(* IEC 61131-3 sources: KinematicsSimulation/crates/sim-opcua/examples/plc/codesys, 3 files *)

(* ---- sim_cycle.st ---- *)
(*
    A PLC cycle against the KinematicsSimulation link (sim-opcua), for CODESYS V3.5 with the CODESYS OPC UA Client
    SL (PLCopen "OPC UA Client for IEC 61131-3" blocks). Uses SIM_Access, SIM_MC_Power and SIM_MC_MoveAbsolute from
    sim_plcopen.st in this folder.

    NOT COMPILED: CODESYS needs a CODESYS Store account to download, so it was not built. The names follow the
    PLCopen specification OPC 30001 (PLCopen-CFB) v1.02, checked 14 November 2026 at reference.opcfoundation.org.
    CHECK: CODESYS's public help shows only its object-oriented "OPC UA Client" library (Client, Read, Write, ...),
    not these PLCopen blocks; a library that offers them may need its namespace prefix. Spec v1.02 also lists
    UA_NamespaceGetIndex, UA_NodeGetHandle, UA_Read and UA_Write as phased out in favour of their *List variants.

    PRG_SimCycle does what ../twincat/sim_cycle.st does: connect with Basic256Sha256 SignAndEncrypt (or None) and
    optionally user name and password, find the namespace index, power the axis, MC_MoveAbsolute, write a path and
    run it, wait until status.busy falls, switch off and disconnect; meanwhile it reads the axis position and
    following error every cycle through node handles got once. Run it in a task of 10 ms.

    Data types (docs/plc.md, "Node ids and data types"): Double -> LREAL, Boolean -> BOOL, UInt16 -> UINT,
    Int32 -> DINT, UInt64 -> ULINT, String -> STRING. The value of UA_Read/UA_Write is an IN_OUT of type ANY: its
    IEC type is what goes on the wire, so it has to be the one in the table.
*)

FUNCTION_BLOCK SIM_CyclicRead
(* Reads one LREAL variable over and over through a node handle that is got once. *)
VAR_INPUT
    xEnable     : BOOL;
    hConnection : DWORD;
    uiNamespace : UINT;
    sNode       : STRING(255);
END_VAR
VAR_OUTPUT
    lrValue   : LREAL;
    udiReads  : UDINT;
    xError    : BOOL;
    dwErrorID : DWORD;
END_VAR
VAR
    fbGetHandle : UA_NodeGetHandle;
    fbRead      : UA_Read;
    fbRelease   : UA_NodeReleaseHandle;
    stNodeID    : UANodeID;
    stInfo      : UANodeAdditionalInfo;
    hNode       : DWORD;
    iStep       : INT;
END_VAR

CASE iStep OF
0:  IF xEnable THEN
        stNodeID.NamespaceIndex := uiNamespace;
        stNodeID.Identifier := sNode;
        stNodeID.IdentifierType := UAIdentifierType.UAIT_String;
        stInfo.AttributeID := 13;   (* the Value attribute *)
        xError := FALSE; dwErrorID := 0;
        iStep := 1;
    END_IF
1:  fbGetHandle(Execute := TRUE, ConnectionHdl := hConnection, NodeID := stNodeID, Timeout := T#5S);
    IF fbGetHandle.Done THEN
        hNode := fbGetHandle.NodeHdl; fbGetHandle(Execute := FALSE, ConnectionHdl := hConnection, NodeID := stNodeID);
        iStep := 2;
    ELSIF fbGetHandle.Error THEN
        dwErrorID := fbGetHandle.ErrorID; fbGetHandle(Execute := FALSE, ConnectionHdl := hConnection, NodeID := stNodeID);
        xError := TRUE; iStep := 9;
    END_IF
2:  (* once a read is done the next starts in the same cycle *)
    fbRead(Execute := TRUE, ConnectionHdl := hConnection, NodeHdl := hNode, NodeAddInfo := stInfo, Timeout := T#5S,
           Variable := lrValue);
    IF fbRead.Done OR fbRead.Error THEN
        IF fbRead.Error THEN xError := TRUE; dwErrorID := fbRead.ErrorID; ELSE udiReads := udiReads + 1; END_IF
        fbRead(Execute := FALSE, Variable := lrValue);
        IF xEnable THEN
            fbRead(Execute := TRUE, ConnectionHdl := hConnection, NodeHdl := hNode, NodeAddInfo := stInfo,
                   Timeout := T#5S, Variable := lrValue);
        ELSE
            iStep := 3;
        END_IF
    END_IF
3:  fbRelease(Execute := TRUE, ConnectionHdl := hConnection, NodeHdl := hNode, Timeout := T#5S);
    IF fbRelease.Done OR fbRelease.Error THEN
        fbRelease(Execute := FALSE, ConnectionHdl := hConnection, NodeHdl := hNode); iStep := 0;
    END_IF
9:  IF NOT xEnable THEN iStep := 0; END_IF
END_CASE
END_FUNCTION_BLOCK

FUNCTION_BLOCK SIM_WriteString
(* One write of a STRING variable: get the handle, write, release. *)
VAR_INPUT
    xExecute    : BOOL;
    hConnection : DWORD;
    uiNamespace : UINT;
    sNode       : STRING(255);
END_VAR
VAR_IN_OUT
    sValue : STRING(255);
END_VAR
VAR_OUTPUT
    xDone : BOOL; xError : BOOL; dwErrorID : DWORD;
END_VAR
VAR
    fbGetHandle : UA_NodeGetHandle;
    fbWrite     : UA_Write;
    fbRelease   : UA_NodeReleaseHandle;
    stNodeID    : UANodeID;
    stInfo      : UANodeAdditionalInfo;
    hNode       : DWORD;
    iStep       : INT;
    xLast       : BOOL;
END_VAR

IF xExecute AND NOT xLast THEN
    xDone := FALSE; xError := FALSE; dwErrorID := 0;
    stNodeID.NamespaceIndex := uiNamespace;
    stNodeID.Identifier := sNode;
    stNodeID.IdentifierType := UAIdentifierType.UAIT_String;
    stInfo.AttributeID := 13;
    iStep := 1;
END_IF
xLast := xExecute;

CASE iStep OF
1:  fbGetHandle(Execute := TRUE, ConnectionHdl := hConnection, NodeID := stNodeID, Timeout := T#5S);
    IF fbGetHandle.Done THEN
        hNode := fbGetHandle.NodeHdl; fbGetHandle(Execute := FALSE, ConnectionHdl := hConnection, NodeID := stNodeID);
        iStep := 2;
    ELSIF fbGetHandle.Error THEN
        dwErrorID := fbGetHandle.ErrorID; fbGetHandle(Execute := FALSE, ConnectionHdl := hConnection, NodeID := stNodeID);
        xError := TRUE; iStep := 0;
    END_IF
2:  fbWrite(Execute := TRUE, ConnectionHdl := hConnection, NodeHdl := hNode, NodeAddInfo := stInfo, Timeout := T#5S,
            Variable := sValue);
    IF fbWrite.Done OR fbWrite.Error THEN
        xError := fbWrite.Error; dwErrorID := fbWrite.ErrorID;
        fbWrite(Execute := FALSE, Variable := sValue);
        iStep := 3;
    END_IF
3:  fbRelease(Execute := TRUE, ConnectionHdl := hConnection, NodeHdl := hNode, Timeout := T#5S);
    IF fbRelease.Done OR fbRelease.Error THEN
        fbRelease(Execute := FALSE, ConnectionHdl := hConnection, NodeHdl := hNode);
        xDone := NOT xError; iStep := 0;
    END_IF
END_CASE
END_FUNCTION_BLOCK

PROGRAM PRG_SimCycle
VAR
    sServerUrl   : STRING(255) := 'opc.tcp://127.0.0.1:4840';   (* sim-opcua on the same PC *)
    xSecure      : BOOL := TRUE;                                 (* FALSE: SecurityPolicy None *)
    sUser        : STRING(63) := '';                             (* empty: anonymous; else as sim-opcua --user *)
    sPassword    : STRING(63) := '';
    sAxis        : STRING(31) := 'x';
    lrTarget     : LREAL := 0.4;
    sPath        : STRING(255) := 'line,0.4,0.25$Nline,0.1,0.25$Nline,0.1,0.35';
    (* FALSE: the position alone, one Read request a cycle, so that status.client_read_* show the task's cycle *)
    xReadFollowingError : BOOL := TRUE;

    fbConnect    : UA_Connect;
    fbNamespace  : UA_NamespaceGetIndex;
    fbDisconnect : UA_Disconnect;
    stSession    : UASessionConnectInfo;
    hConnection  : DWORD;
    uiNamespace  : UINT;
    fbPower      : SIM_MC_Power;
    fbMove       : SIM_MC_MoveAbsolute;
    fbPath       : SIM_WriteString;
    fbAccess     : SIM_Access;
    fbPosition   : SIM_CyclicRead;
    fbError      : SIM_CyclicRead;
    xFlag        : BOOL;
    lrUnused     : LREAL;
    uiUnused     : UINT;
    xBusySeen    : BOOL;
    lrLargestError : LREAL;
    iStep        : INT;
END_VAR

CASE iStep OF
0:  stSession.ApplicationName := 'CODESYS sim client';
    IF xSecure THEN
        (* The client certificate: create it in View > Security Screen, Devices tab, for the device. sim-opcua
           refuses it once and stores it in pki/rejected; move it to pki/trusted, or run sim-opcua with --trust-all
           while commissioning. The server's certificate (pki/own/cert.der) lands in the device's "Certificates in
           Quarantine" on the first attempt: drag it to "Trusted Certificates" in the same tab. *)
        stSession.SecurityMsgMode := UASecurityMsgMode.UASMM_SignEncrypt;
        stSession.SecurityPolicy := UASecurityPolicy.UASP_Basic256Sha256;
    ELSE
        stSession.SecurityMsgMode := UASecurityMsgMode.UASMM_None;
        stSession.SecurityPolicy := UASecurityPolicy.UASP_None;
    END_IF
    IF LEN(sUser) > 0 THEN
        stSession.UserIdentityToken.UserIdentityTokenType := UAUserIdentityTokenType.UAUITT_Username;
        stSession.UserIdentityToken.TokenParam1 := sUser;
        stSession.UserIdentityToken.TokenParam2 := sPassword;
    END_IF
    fbConnect(Execute := TRUE, ServerEndpointUrl := sServerUrl, SessionConnectInfo := stSession, Timeout := T#5S);
    IF fbConnect.Done THEN hConnection := fbConnect.ConnectionHdl; fbConnect(Execute := FALSE); iStep := 10;
    ELSIF fbConnect.Error THEN fbConnect(Execute := FALSE); iStep := 900; END_IF
10: fbNamespace(Execute := TRUE, ConnectionHdl := hConnection, NamespaceUri := 'urn:kinematics-simulation', Timeout := T#5S);
    IF fbNamespace.Done THEN uiNamespace := fbNamespace.NamespaceIndex; fbNamespace(Execute := FALSE); iStep := 20;
    ELSIF fbNamespace.Error THEN fbNamespace(Execute := FALSE); iStep := 900; END_IF
20: fbPower.Enable := TRUE;
    IF fbPower.Status THEN iStep := 30; END_IF
30: fbMove.Position := lrTarget; fbMove.Velocity := 0.5; fbMove.Acceleration := 5.0; fbMove.Deceleration := 5.0;
    fbMove.Jerk := 100.0;
    fbMove.Execute := TRUE;
    IF fbMove.Done THEN fbMove.Execute := FALSE; iStep := 40;
    ELSIF fbMove.Error OR fbMove.CommandAborted THEN iStep := 900; END_IF
40: fbPath(xExecute := FALSE, sValue := sPath);
    fbPath(xExecute := TRUE, hConnection := hConnection, uiNamespace := uiNamespace, sNode := 'command.path', sValue := sPath);
    IF fbPath.xDone THEN iStep := 42; ELSIF fbPath.xError THEN iStep := 900; ELSE iStep := 41; END_IF
41: fbPath(xExecute := TRUE, sValue := sPath);
    IF fbPath.xDone THEN iStep := 42; ELSIF fbPath.xError THEN iStep := 900; END_IF
42: xFlag := TRUE;
    fbAccess(xExecute := FALSE, xValue := xFlag, lrValue := lrUnused, uiValue := uiUnused);
    fbAccess(xExecute := TRUE, hConnection := hConnection, uiNamespace := uiNamespace, sNode := 'command.run_path',
             eKind := SIM_BOOL, xWrite := TRUE, xValue := xFlag, lrValue := lrUnused, uiValue := uiUnused);
    iStep := 43;
43: fbAccess(xExecute := TRUE, xValue := xFlag, lrValue := lrUnused, uiValue := uiUnused);
    IF fbAccess.xDone THEN xBusySeen := FALSE; iStep := 50; ELSIF fbAccess.xError THEN iStep := 900; END_IF
50: (* poll status.busy until the path is over *)
    fbAccess(xExecute := FALSE, xValue := xFlag, lrValue := lrUnused, uiValue := uiUnused);
    fbAccess(xExecute := TRUE, hConnection := hConnection, uiNamespace := uiNamespace, sNode := 'status.busy',
             eKind := SIM_BOOL, xWrite := FALSE, xValue := xFlag, lrValue := lrUnused, uiValue := uiUnused);
    iStep := 51;
51: fbAccess(xExecute := TRUE, xValue := xFlag, lrValue := lrUnused, uiValue := uiUnused);
    IF fbAccess.xDone THEN
        IF xFlag THEN xBusySeen := TRUE; iStep := 50;
        ELSIF xBusySeen THEN iStep := 60;
        ELSE iStep := 50; END_IF
    ELSIF fbAccess.xError THEN iStep := 900; END_IF
60: fbPower.Enable := FALSE;
    IF NOT fbPower.Status THEN iStep := 70; END_IF
70: fbDisconnect(Execute := TRUE, ConnectionHdl := hConnection, Timeout := T#5S);
    IF fbDisconnect.Done OR fbDisconnect.Error THEN fbDisconnect(Execute := FALSE); iStep := 100; END_IF
100: ; (* finished: lrLargestError holds the largest following error *)
900: ; (* error: look at the blocks' ErrorID and at status.refused on the server *)
END_CASE

fbPosition(xEnable := iStep >= 20 AND iStep < 70, hConnection := hConnection, uiNamespace := uiNamespace,
           sNode := CONCAT(CONCAT('signal.axis.', sAxis), '.position'));
fbError(xEnable := xReadFollowingError AND iStep >= 20 AND iStep < 70, hConnection := hConnection, uiNamespace := uiNamespace,
        sNode := CONCAT(CONCAT('signal.axis.', sAxis), '.following_error'));
IF ABS(fbError.lrValue) > lrLargestError THEN lrLargestError := ABS(fbError.lrValue); END_IF

IF iStep >= 20 AND iStep < 70 THEN
    fbPower(hConnection := hConnection, uiNamespace := uiNamespace, sAxis := sAxis);
    fbMove(hConnection := hConnection, uiNamespace := uiNamespace, sAxis := sAxis);
END_IF
END_PROGRAM

(* ---- sim_plcopen.st ---- *)
(*
    PLCopen motion over OPC UA to the KinematicsSimulation link (sim-opcua), for CODESYS V3.5.
    Library: CODESYS OPC UA Client SL (the PLCopen "OPC UA Client for IEC 61131-3" function blocks UA_Connect,
    UA_NamespaceGetIndex, UA_NodeGetHandle, UA_Read, UA_Write, UA_NodeReleaseHandle, UA_Disconnect).

    NOT COMPILED: CODESYS needs a CODESYS Store account to download, so this file was not built. The names follow
    the PLCopen specification OPC 30001 (PLCopen-CFB) v1.02, checked 14 November 2026 at
    reference.opcfoundation.org. CHECK: CODESYS's public help shows only its object-oriented "OPC UA Client"
    library, not these PLCopen blocks; a library that offers them may need its namespace prefix. Spec v1.02 lists
    UA_NamespaceGetIndex, UA_NodeGetHandle, UA_Read and UA_Write as phased out in favour of their *List variants.

    The structure is the one of ../twincat/sim_plcopen.st. The PLCopen UA_Read and UA_Write take the value as
    VAR_IN_OUT of type ANY, so SIM_Access keeps one buffer per data type instead of a pointer.
*)

TYPE E_SimKind : (SIM_BOOL, SIM_LREAL, SIM_UINT); END_TYPE

FUNCTION_BLOCK SIM_Access
VAR_INPUT
    xExecute    : BOOL;
    hConnection : DWORD;
    uiNamespace : UINT;
    sNode       : STRING(255);
    eKind       : E_SimKind;
    xWrite      : BOOL;     (* TRUE: write the value below; FALSE: read into it *)
END_VAR
VAR_IN_OUT
    xValue  : BOOL;
    lrValue : LREAL;
    uiValue : UINT;
END_VAR
VAR_OUTPUT
    xDone    : BOOL;
    xBusy    : BOOL;
    xError   : BOOL;
    dwErrorID : DWORD;
END_VAR
VAR
    fbGetHandle : UA_NodeGetHandle;
    fbReadBool, fbReadReal, fbReadUint    : UA_Read;
    fbWriteBool, fbWriteReal, fbWriteUint : UA_Write;
    fbRelease   : UA_NodeReleaseHandle;
    stNodeID    : UANodeID;
    stInfo      : UANodeAdditionalInfo;
    hNode       : DWORD;
    iStep       : INT;
    xLast       : BOOL;
    xAccessDone, xAccessError : BOOL;
    dwAccessError : DWORD;
END_VAR

IF xExecute AND NOT xLast THEN
    xDone := FALSE; xError := FALSE; dwErrorID := 0; xBusy := TRUE;
    stNodeID.NamespaceIndex := uiNamespace;
    stNodeID.Identifier := sNode;
    stNodeID.IdentifierType := UAIdentifierType.UAIT_String;
    stInfo.AttributeID := 13;   (* the Value attribute *)
    iStep := 1;
END_IF
xLast := xExecute;

CASE iStep OF
1:  fbGetHandle(Execute := TRUE, ConnectionHdl := hConnection, NodeID := stNodeID, Timeout := T#5S);
    IF fbGetHandle.Done THEN
        hNode := fbGetHandle.NodeHdl;
        fbGetHandle(Execute := FALSE, ConnectionHdl := hConnection, NodeID := stNodeID);
        iStep := 2;
    ELSIF fbGetHandle.Error THEN
        dwErrorID := fbGetHandle.ErrorID;
        fbGetHandle(Execute := FALSE, ConnectionHdl := hConnection, NodeID := stNodeID);
        xError := TRUE; xBusy := FALSE; iStep := 0;
    END_IF
2:  (* one instance per data type, because the value is an IN_OUT of type ANY *)
    CASE eKind OF
    SIM_BOOL:
        IF xWrite THEN
            fbWriteBool(Execute := TRUE, ConnectionHdl := hConnection, NodeHdl := hNode, NodeAddInfo := stInfo, Timeout := T#5S, Variable := xValue);
            xAccessDone := fbWriteBool.Done; xAccessError := fbWriteBool.Error; dwAccessError := fbWriteBool.ErrorID;
            IF xAccessDone OR xAccessError THEN fbWriteBool(Execute := FALSE, Variable := xValue); END_IF
        ELSE
            fbReadBool(Execute := TRUE, ConnectionHdl := hConnection, NodeHdl := hNode, NodeAddInfo := stInfo, Timeout := T#5S, Variable := xValue);
            xAccessDone := fbReadBool.Done; xAccessError := fbReadBool.Error; dwAccessError := fbReadBool.ErrorID;
            IF xAccessDone OR xAccessError THEN fbReadBool(Execute := FALSE, Variable := xValue); END_IF
        END_IF
    SIM_LREAL:
        IF xWrite THEN
            fbWriteReal(Execute := TRUE, ConnectionHdl := hConnection, NodeHdl := hNode, NodeAddInfo := stInfo, Timeout := T#5S, Variable := lrValue);
            xAccessDone := fbWriteReal.Done; xAccessError := fbWriteReal.Error; dwAccessError := fbWriteReal.ErrorID;
            IF xAccessDone OR xAccessError THEN fbWriteReal(Execute := FALSE, Variable := lrValue); END_IF
        ELSE
            fbReadReal(Execute := TRUE, ConnectionHdl := hConnection, NodeHdl := hNode, NodeAddInfo := stInfo, Timeout := T#5S, Variable := lrValue);
            xAccessDone := fbReadReal.Done; xAccessError := fbReadReal.Error; dwAccessError := fbReadReal.ErrorID;
            IF xAccessDone OR xAccessError THEN fbReadReal(Execute := FALSE, Variable := lrValue); END_IF
        END_IF
    SIM_UINT:
        IF xWrite THEN
            fbWriteUint(Execute := TRUE, ConnectionHdl := hConnection, NodeHdl := hNode, NodeAddInfo := stInfo, Timeout := T#5S, Variable := uiValue);
            xAccessDone := fbWriteUint.Done; xAccessError := fbWriteUint.Error; dwAccessError := fbWriteUint.ErrorID;
            IF xAccessDone OR xAccessError THEN fbWriteUint(Execute := FALSE, Variable := uiValue); END_IF
        ELSE
            fbReadUint(Execute := TRUE, ConnectionHdl := hConnection, NodeHdl := hNode, NodeAddInfo := stInfo, Timeout := T#5S, Variable := uiValue);
            xAccessDone := fbReadUint.Done; xAccessError := fbReadUint.Error; dwAccessError := fbReadUint.ErrorID;
            IF xAccessDone OR xAccessError THEN fbReadUint(Execute := FALSE, Variable := uiValue); END_IF
        END_IF
    END_CASE
    IF xAccessDone OR xAccessError THEN
        xError := xAccessError; dwErrorID := dwAccessError;
        iStep := 3;
    END_IF
3:  fbRelease(Execute := TRUE, ConnectionHdl := hConnection, NodeHdl := hNode, Timeout := T#5S);
    IF fbRelease.Done OR fbRelease.Error THEN
        fbRelease(Execute := FALSE, ConnectionHdl := hConnection, NodeHdl := hNode);
        xBusy := FALSE; xDone := NOT xError; iStep := 0;
    END_IF
END_CASE
END_FUNCTION_BLOCK

FUNCTION_BLOCK SIM_Handshake
VAR_INPUT
    Execute     : BOOL;
    hConnection : DWORD;
    uiNamespace : UINT;
    sAxis       : STRING(31);
    sFb         : STRING(31);                  (* 'Home', 'MoveAbsolute', 'MoveRelative', 'Stop', 'Reset' *)
    iParams     : INT;                         (* 0..5 *)
    asParam     : ARRAY[1..5] OF STRING(31);
    alrParam    : ARRAY[1..5] OF LREAL;
END_VAR
VAR_OUTPUT
    Done           : BOOL;
    Busy           : BOOL;
    Active         : BOOL;
    CommandAborted : BOOL;
    Error          : BOOL;
    ErrorID        : UINT;
END_VAR
VAR
    fbAccess : SIM_Access;
    iPhase   : INT;      (* 0 idle, 1 inputs, 2 Execute low, 3 wait Done low, 4 Execute high, 5 poll, 6 finished *)
    iItem    : INT;
    xLast    : BOOL;
    xStarted : BOOL;
    xValue   : BOOL;
    lrValue  : LREAL;
    uiValue  : UINT;
    axRemote : ARRAY[1..4] OF BOOL;   (* Busy, Done, CommandAborted, Error as read *)
    sBase    : STRING(80);
END_VAR

IF Execute AND NOT xLast THEN
    Done := FALSE; Busy := TRUE; Active := FALSE; CommandAborted := FALSE; Error := FALSE; ErrorID := 0;
    sBase := CONCAT(CONCAT(CONCAT('axis.', sAxis), '.'), CONCAT(sFb, '.'));
    IF iParams > 0 THEN iPhase := 1; ELSE iPhase := 2; END_IF
    iItem := 1; xStarted := FALSE;
ELSIF NOT Execute AND xLast THEN
    Done := FALSE; CommandAborted := FALSE; Error := FALSE; ErrorID := 0;
    IF NOT Busy THEN iPhase := 2; iItem := 1; xStarted := FALSE; END_IF
END_IF
xLast := Execute;

IF iPhase > 0 AND iPhase < 6 THEN
    IF NOT xStarted THEN
        CASE iPhase OF
        1:  fbAccess.sNode := CONCAT(sBase, asParam[iItem]); lrValue := alrParam[iItem];
            fbAccess.eKind := SIM_LREAL; fbAccess.xWrite := TRUE;
        2, 4:
            fbAccess.sNode := CONCAT(sBase, 'Execute'); xValue := iPhase = 4;
            fbAccess.eKind := SIM_BOOL; fbAccess.xWrite := TRUE;
        3:  fbAccess.sNode := CONCAT(sBase, 'Done');
            fbAccess.eKind := SIM_BOOL; fbAccess.xWrite := FALSE;
        5:  CASE iItem OF
            1: fbAccess.sNode := CONCAT(sBase, 'Busy');
            2: fbAccess.sNode := CONCAT(sBase, 'Done');
            3: fbAccess.sNode := CONCAT(sBase, 'CommandAborted');
            4: fbAccess.sNode := CONCAT(sBase, 'Error');
            ELSE fbAccess.sNode := CONCAT(sBase, 'ErrorID');
            END_CASE
            IF iItem <= 4 THEN fbAccess.eKind := SIM_BOOL; ELSE fbAccess.eKind := SIM_UINT; END_IF
            fbAccess.xWrite := FALSE;
        END_CASE
        fbAccess(xExecute := FALSE, hConnection := hConnection, uiNamespace := uiNamespace, xValue := xValue, lrValue := lrValue, uiValue := uiValue);
        xStarted := TRUE;
    END_IF
    fbAccess(xExecute := TRUE, hConnection := hConnection, uiNamespace := uiNamespace, xValue := xValue, lrValue := lrValue, uiValue := uiValue);

    IF fbAccess.xError THEN
        Error := TRUE; ErrorID := 16#FFFF; Busy := FALSE; iPhase := 6;   (* the OPC UA access failed *)
    ELSIF fbAccess.xDone THEN
        xStarted := FALSE;
        CASE iPhase OF
        1:  iItem := iItem + 1;
            IF iItem > iParams THEN iPhase := 2; iItem := 1; END_IF
        2:  IF Busy THEN iPhase := 3; ELSE iPhase := 0; END_IF
        3:  IF NOT xValue THEN iPhase := 4; END_IF   (* outputs are published once a cycle *)
        4:  iPhase := 5; iItem := 1;
        5:  IF iItem <= 4 THEN
                axRemote[iItem] := xValue;
                iItem := iItem + 1;
            ELSE
                ErrorID := uiValue;
                Active := axRemote[1];
                IF axRemote[2] OR axRemote[3] OR axRemote[4] THEN
                    Done := axRemote[2] AND Execute;
                    CommandAborted := axRemote[3] AND Execute;
                    Error := axRemote[4] AND Execute;
                    Busy := FALSE; Active := FALSE;
                    iPhase := 6;
                END_IF
                iItem := 1;
            END_IF
        END_CASE
    END_IF
END_IF
END_FUNCTION_BLOCK

FUNCTION_BLOCK SIM_MC_Power
VAR_INPUT
    Enable : BOOL; hConnection : DWORD; uiNamespace : UINT; sAxis : STRING(31);
END_VAR
VAR_OUTPUT
    Status : BOOL; Valid : BOOL; Error : BOOL;
END_VAR
VAR
    fbAccess : SIM_Access;
    iStep    : INT;
    xWritten : BOOL;
    xFirst   : BOOL := TRUE;
    xValue   : BOOL;
    lrDummy  : LREAL;
    uiDummy  : UINT;
END_VAR

(* writes Enable when it changes, otherwise reads Power.Status *)
IF iStep = 0 THEN
    fbAccess.eKind := SIM_BOOL;
    IF xFirst OR Enable <> xWritten THEN
        xValue := Enable; xWritten := Enable; xFirst := FALSE;
        fbAccess.sNode := CONCAT(CONCAT('axis.', sAxis), '.Power.Enable'); fbAccess.xWrite := TRUE;
    ELSE
        fbAccess.sNode := CONCAT(CONCAT('axis.', sAxis), '.Power.Status'); fbAccess.xWrite := FALSE;
    END_IF
    fbAccess(xExecute := FALSE, hConnection := hConnection, uiNamespace := uiNamespace, xValue := xValue, lrValue := lrDummy, uiValue := uiDummy);
    iStep := 1;
END_IF
fbAccess(xExecute := TRUE, hConnection := hConnection, uiNamespace := uiNamespace, xValue := xValue, lrValue := lrDummy, uiValue := uiDummy);
IF fbAccess.xDone OR fbAccess.xError THEN
    Error := fbAccess.xError;
    IF fbAccess.xDone AND NOT fbAccess.xWrite THEN Status := xValue; END_IF
    Valid := Status AND NOT Error;
    iStep := 0;
END_IF
END_FUNCTION_BLOCK

FUNCTION_BLOCK SIM_MC_Home
VAR_INPUT
    Execute : BOOL; hConnection : DWORD; uiNamespace : UINT; sAxis : STRING(31);
END_VAR
VAR_OUTPUT
    Done : BOOL; Busy : BOOL; Active : BOOL; CommandAborted : BOOL; Error : BOOL; ErrorID : UINT;
END_VAR
VAR
    fbCall : SIM_Handshake;
END_VAR
fbCall(Execute := Execute, hConnection := hConnection, uiNamespace := uiNamespace, sAxis := sAxis, sFb := 'Home', iParams := 0);
Done := fbCall.Done; Busy := fbCall.Busy; Active := fbCall.Active;
CommandAborted := fbCall.CommandAborted; Error := fbCall.Error; ErrorID := fbCall.ErrorID;
END_FUNCTION_BLOCK

FUNCTION_BLOCK SIM_MC_MoveAbsolute
VAR_INPUT
    Execute : BOOL; hConnection : DWORD; uiNamespace : UINT; sAxis : STRING(31);
    Position : LREAL; Velocity : LREAL; Acceleration : LREAL; Deceleration : LREAL; Jerk : LREAL;
END_VAR
VAR_OUTPUT
    Done : BOOL; Busy : BOOL; Active : BOOL; CommandAborted : BOOL; Error : BOOL; ErrorID : UINT;
END_VAR
VAR
    fbCall : SIM_Handshake;
END_VAR
fbCall.asParam[1] := 'Position';     fbCall.alrParam[1] := Position;
fbCall.asParam[2] := 'Velocity';     fbCall.alrParam[2] := Velocity;
fbCall.asParam[3] := 'Acceleration'; fbCall.alrParam[3] := Acceleration;
fbCall.asParam[4] := 'Deceleration'; fbCall.alrParam[4] := Deceleration;
fbCall.asParam[5] := 'Jerk';         fbCall.alrParam[5] := Jerk;
fbCall(Execute := Execute, hConnection := hConnection, uiNamespace := uiNamespace, sAxis := sAxis, sFb := 'MoveAbsolute', iParams := 5);
Done := fbCall.Done; Busy := fbCall.Busy; Active := fbCall.Active;
CommandAborted := fbCall.CommandAborted; Error := fbCall.Error; ErrorID := fbCall.ErrorID;
END_FUNCTION_BLOCK

FUNCTION_BLOCK SIM_MC_MoveRelative
VAR_INPUT
    Execute : BOOL; hConnection : DWORD; uiNamespace : UINT; sAxis : STRING(31);
    Distance : LREAL; Velocity : LREAL; Acceleration : LREAL; Deceleration : LREAL; Jerk : LREAL;
END_VAR
VAR_OUTPUT
    Done : BOOL; Busy : BOOL; Active : BOOL; CommandAborted : BOOL; Error : BOOL; ErrorID : UINT;
END_VAR
VAR
    fbCall : SIM_Handshake;
END_VAR
fbCall.asParam[1] := 'Distance';     fbCall.alrParam[1] := Distance;
fbCall.asParam[2] := 'Velocity';     fbCall.alrParam[2] := Velocity;
fbCall.asParam[3] := 'Acceleration'; fbCall.alrParam[3] := Acceleration;
fbCall.asParam[4] := 'Deceleration'; fbCall.alrParam[4] := Deceleration;
fbCall.asParam[5] := 'Jerk';         fbCall.alrParam[5] := Jerk;
fbCall(Execute := Execute, hConnection := hConnection, uiNamespace := uiNamespace, sAxis := sAxis, sFb := 'MoveRelative', iParams := 5);
Done := fbCall.Done; Busy := fbCall.Busy; Active := fbCall.Active;
CommandAborted := fbCall.CommandAborted; Error := fbCall.Error; ErrorID := fbCall.ErrorID;
END_FUNCTION_BLOCK

FUNCTION_BLOCK SIM_MC_Stop
VAR_INPUT
    Execute : BOOL; hConnection : DWORD; uiNamespace : UINT; sAxis : STRING(31);
    Deceleration : LREAL;
END_VAR
VAR_OUTPUT
    Done : BOOL; Busy : BOOL; Active : BOOL; CommandAborted : BOOL; Error : BOOL; ErrorID : UINT;
END_VAR
VAR
    fbCall : SIM_Handshake;
END_VAR
fbCall.asParam[1] := 'Deceleration'; fbCall.alrParam[1] := Deceleration;
fbCall(Execute := Execute, hConnection := hConnection, uiNamespace := uiNamespace, sAxis := sAxis, sFb := 'Stop', iParams := 1);
Done := fbCall.Done; Busy := fbCall.Busy; Active := fbCall.Active;
CommandAborted := fbCall.CommandAborted; Error := fbCall.Error; ErrorID := fbCall.ErrorID;
END_FUNCTION_BLOCK

FUNCTION_BLOCK SIM_MC_Reset
VAR_INPUT
    Execute : BOOL; hConnection : DWORD; uiNamespace : UINT; sAxis : STRING(31);
END_VAR
VAR_OUTPUT
    Done : BOOL; Busy : BOOL; Error : BOOL; ErrorID : UINT;
END_VAR
VAR
    fbCall : SIM_Handshake;
END_VAR
fbCall(Execute := Execute, hConnection := hConnection, uiNamespace := uiNamespace, sAxis := sAxis, sFb := 'Reset', iParams := 0);
Done := fbCall.Done; Busy := fbCall.Busy; Error := fbCall.Error; ErrorID := fbCall.ErrorID;
END_FUNCTION_BLOCK

PROGRAM PRG_SimDemo
VAR
    fbConnect    : UA_Connect;
    fbNamespace  : UA_NamespaceGetIndex;
    fbDisconnect : UA_Disconnect;
    stSession    : UASessionConnectInfo;
    hConnection  : DWORD;
    uiNamespace  : UINT;
    fbPower      : SIM_MC_Power;
    fbHome       : SIM_MC_Home;
    fbMove       : SIM_MC_MoveAbsolute;
    fbStop       : SIM_MC_Stop;
    tonMoving    : TON;
    iStep        : INT;
    sAxis        : STRING(31) := 'x';
END_VAR

CASE iStep OF
0:  stSession.ApplicationName := 'CODESYS sim client';
    stSession.SecurityMsgMode := UASecurityMsgMode.UASMM_None;
    stSession.SecurityPolicy := UASecurityPolicy.UASP_None;
    fbConnect(Execute := TRUE, ServerEndpointUrl := 'opc.tcp://192.168.0.10:4840', SessionConnectInfo := stSession, Timeout := T#5S);
    IF fbConnect.Done THEN hConnection := fbConnect.ConnectionHdl; fbConnect(Execute := FALSE); iStep := 10;
    ELSIF fbConnect.Error THEN fbConnect(Execute := FALSE); iStep := 900; END_IF
10: fbNamespace(Execute := TRUE, ConnectionHdl := hConnection, NamespaceUri := 'urn:kinematics-simulation', Timeout := T#5S);
    IF fbNamespace.Done THEN uiNamespace := fbNamespace.NamespaceIndex; fbNamespace(Execute := FALSE); iStep := 20;
    ELSIF fbNamespace.Error THEN fbNamespace(Execute := FALSE); iStep := 900; END_IF
20: fbPower.Enable := TRUE;
    IF fbPower.Status THEN iStep := 30; END_IF
30: fbHome.Execute := TRUE;
    IF fbHome.Done THEN fbHome.Execute := FALSE; iStep := 40;
    ELSIF fbHome.Error THEN iStep := 900; END_IF
40: fbMove.Position := 0.6; fbMove.Velocity := 0.5; fbMove.Acceleration := 5.0; fbMove.Deceleration := 5.0; fbMove.Jerk := 100.0;
    fbMove.Execute := TRUE;
    tonMoving(IN := fbMove.Busy, PT := T#500MS);
    IF tonMoving.Q OR fbMove.Done THEN iStep := 50;
    ELSIF fbMove.Error THEN iStep := 900; END_IF
50: fbStop.Deceleration := 2.0;
    fbStop.Execute := TRUE;
    IF fbStop.Done THEN fbStop.Execute := FALSE; fbMove.Execute := FALSE; iStep := 60;
    ELSIF fbStop.Error THEN iStep := 900; END_IF
60: fbPower.Enable := FALSE;
    IF NOT fbPower.Status THEN iStep := 70; END_IF
70: fbDisconnect(Execute := TRUE, ConnectionHdl := hConnection, Timeout := T#5S);
    IF fbDisconnect.Done OR fbDisconnect.Error THEN fbDisconnect(Execute := FALSE); iStep := 100; END_IF
100: ;
900: ;
END_CASE

IF iStep >= 20 AND iStep < 70 THEN
    fbPower(hConnection := hConnection, uiNamespace := uiNamespace, sAxis := sAxis);
    fbHome(hConnection := hConnection, uiNamespace := uiNamespace, sAxis := sAxis);
    fbMove(hConnection := hConnection, uiNamespace := uiNamespace, sAxis := sAxis);
    fbStop(hConnection := hConnection, uiNamespace := uiNamespace, sAxis := sAxis);
END_IF
END_PROGRAM

(* ---- sim_sync.st ---- *)
(*
    PLCopen synchronised motion over OPC UA to the KinematicsSimulation link (sim-opcua), for CODESYS V3.5:
    MC_GearIn, MC_GearOut, MC_CamIn and MC_CamOut on a slave axis, its master another axis of the machine.
    Needs SIM_Access and SIM_Handshake from sim_plcopen.st and SIM_WriteString from sim_cycle.st in the same project.

    NOT COMPILED, as sim_plcopen.st (see its header for the library and the names). It uses only the blocks of
    sim_plcopen.st and sim_cycle.st and plain IEC 61131-3. SIM_WriteString writes a STRING(255): a cam table
    (CamIn.Table) longer than that needs a longer STRING there.

    The structure is the one of ../twincat/sim_sync.st:
      SIM_SyncHandshake    the handshake of MC_GearIn or MC_CamIn: inputs and texts, Execute low, Execute high, then
                           poll Busy, InGear/InSync, CommandAborted, Error and ErrorID for as long as the block is busy:
                           unlike a move it stays busy while the slave is coupled
      SIM_MC_GearIn, SIM_MC_CamIn, SIM_MC_GearOut, SIM_MC_CamOut   thin wrappers with PLCopen inputs and outputs
      PRG_SimSyncDemo      x moves, y gears in at 2:1, gears out, cams in on a 3-4-5 table, cams out, stops
*)

FUNCTION_BLOCK SIM_SyncHandshake
VAR_INPUT
    Execute     : BOOL;
    hConnection : DWORD;
    uiNamespace : UINT;
    sAxis       : STRING(31);                  (* the slave's axis id *)
    sFb         : STRING(31);                  (* 'GearIn' or 'CamIn' *)
    sMaster     : STRING(31);                  (* the master's axis id; '' for the machine's virtual cam master *)
    sTable      : STRING(255);                 (* CamIn only: the cam table, '' to leave it as it is *)
    iParams     : INT;                         (* 0..6 *)
    asParam     : ARRAY[1..6] OF STRING(31);
    alrParam    : ARRAY[1..6] OF LREAL;
END_VAR
VAR_OUTPUT
    InSync         : BOOL;     (* InGear of MC_GearIn, InSync of MC_CamIn *)
    Busy           : BOOL;
    Active         : BOOL;
    CommandAborted : BOOL;
    Error          : BOOL;
    ErrorID        : UINT;
END_VAR
VAR
    fbAccess : SIM_Access;
    fbText   : SIM_WriteString;
    iPhase   : INT;      (* 0 idle, 1 inputs, 2 Master, 3 Table, 4 Execute low, 5 Execute high, 6 poll, 7 finished *)
    iItem    : INT;
    xLast    : BOOL;
    xStarted : BOOL;
    xValue   : BOOL;
    lrValue  : LREAL;
    uiValue  : UINT;
    sText    : STRING(255);
    axRemote : ARRAY[1..4] OF BOOL;   (* Busy, InGear/InSync, CommandAborted, Error as read *)
    sBase    : STRING(80);
    sSync    : STRING(31);
END_VAR

IF Execute AND NOT xLast THEN
    InSync := FALSE; Busy := TRUE; Active := FALSE; CommandAborted := FALSE; Error := FALSE; ErrorID := 0;
    sBase := CONCAT(CONCAT(CONCAT('axis.', sAxis), '.'), CONCAT(sFb, '.'));
    IF sFb = 'GearIn' THEN sSync := 'InGear'; ELSE sSync := 'InSync'; END_IF
    IF iParams > 0 THEN iPhase := 1; ELSE iPhase := 2; END_IF
    iItem := 1; xStarted := FALSE;
ELSIF NOT Execute AND xLast THEN
    (* the outputs fall with Execute; a coupled block stays coupled until GearOut/CamOut or another block *)
    InSync := FALSE; CommandAborted := FALSE; Error := FALSE; ErrorID := 0;
    iPhase := 4; xStarted := FALSE;
END_IF
xLast := Execute;

IF iPhase = 2 OR iPhase = 3 THEN
    (* the texts: the master, then (CamIn) the table *)
    IF iPhase = 3 AND (sFb <> 'CamIn' OR LEN(sTable) = 0) THEN
        iPhase := 4;
    ELSE
        IF NOT xStarted THEN
            IF iPhase = 2 THEN
                fbText.sNode := CONCAT(sBase, 'Master'); sText := sMaster;
            ELSE
                fbText.sNode := CONCAT(sBase, 'Table'); sText := sTable;
            END_IF
            fbText(xExecute := FALSE, hConnection := hConnection, uiNamespace := uiNamespace, sValue := sText);
            xStarted := TRUE;
        END_IF
        fbText(xExecute := TRUE, hConnection := hConnection, uiNamespace := uiNamespace, sValue := sText);
        IF fbText.xError THEN
            Error := TRUE; ErrorID := 16#FFFF; Busy := FALSE; iPhase := 7;
        ELSIF fbText.xDone THEN
            xStarted := FALSE; iPhase := iPhase + 1;
        END_IF
    END_IF
ELSIF iPhase > 0 AND iPhase < 7 THEN
    IF NOT xStarted THEN
        CASE iPhase OF
        1:  fbAccess.sNode := CONCAT(sBase, asParam[iItem]); lrValue := alrParam[iItem];
            fbAccess.eKind := SIM_LREAL; fbAccess.xWrite := TRUE;
        4, 5:
            fbAccess.sNode := CONCAT(sBase, 'Execute'); xValue := iPhase = 5 AND Execute;
            fbAccess.eKind := SIM_BOOL; fbAccess.xWrite := TRUE;
        6:  CASE iItem OF
            1: fbAccess.sNode := CONCAT(sBase, 'Busy');
            2: fbAccess.sNode := CONCAT(sBase, sSync);
            3: fbAccess.sNode := CONCAT(sBase, 'CommandAborted');
            4: fbAccess.sNode := CONCAT(sBase, 'Error');
            ELSE fbAccess.sNode := CONCAT(sBase, 'ErrorID');
            END_CASE
            IF iItem <= 4 THEN fbAccess.eKind := SIM_BOOL; ELSE fbAccess.eKind := SIM_UINT; END_IF
            fbAccess.xWrite := FALSE;
        END_CASE
        fbAccess(xExecute := FALSE, hConnection := hConnection, uiNamespace := uiNamespace, xValue := xValue, lrValue := lrValue, uiValue := uiValue);
        xStarted := TRUE;
    END_IF
    fbAccess(xExecute := TRUE, hConnection := hConnection, uiNamespace := uiNamespace, xValue := xValue, lrValue := lrValue, uiValue := uiValue);

    IF fbAccess.xError THEN
        Error := TRUE; ErrorID := 16#FFFF; Busy := FALSE; iPhase := 7;   (* the OPC UA access failed *)
    ELSIF fbAccess.xDone THEN
        xStarted := FALSE;
        CASE iPhase OF
        1:  iItem := iItem + 1;
            IF iItem > iParams THEN iPhase := 2; iItem := 1; END_IF
        4:  IF Execute THEN iPhase := 5; ELSE iPhase := 0; Busy := FALSE; Active := FALSE; END_IF
        5:  iPhase := 6; iItem := 1;
        6:  IF iItem <= 4 THEN
                axRemote[iItem] := xValue;
                iItem := iItem + 1;
            ELSE
                ErrorID := uiValue;
                Busy := axRemote[1]; Active := axRemote[1];
                InSync := axRemote[2] AND Execute;
                CommandAborted := axRemote[3] AND Execute;
                Error := axRemote[4] AND Execute;
                (* coupled, the block stays busy: poll on; it is over once it is no longer busy *)
                IF NOT Busy THEN iPhase := 7; END_IF
                iItem := 1;
            END_IF
        END_CASE
    END_IF
END_IF
END_FUNCTION_BLOCK

FUNCTION_BLOCK SIM_MC_GearIn
VAR_INPUT
    Execute : BOOL; hConnection : DWORD; uiNamespace : UINT;
    sMaster : STRING(31); sSlave : STRING(31);
    RatioNumerator : LREAL; RatioDenominator : LREAL; Acceleration : LREAL; Deceleration : LREAL; Jerk : LREAL;
END_VAR
VAR_OUTPUT
    InGear : BOOL; Busy : BOOL; Active : BOOL; CommandAborted : BOOL; Error : BOOL; ErrorID : UINT;
END_VAR
VAR
    fbCall : SIM_SyncHandshake;
END_VAR
fbCall.asParam[1] := 'RatioNumerator';   fbCall.alrParam[1] := RatioNumerator;
fbCall.asParam[2] := 'RatioDenominator'; fbCall.alrParam[2] := RatioDenominator;
fbCall.asParam[3] := 'Acceleration';     fbCall.alrParam[3] := Acceleration;
fbCall.asParam[4] := 'Deceleration';     fbCall.alrParam[4] := Deceleration;
fbCall.asParam[5] := 'Jerk';             fbCall.alrParam[5] := Jerk;
fbCall(Execute := Execute, hConnection := hConnection, uiNamespace := uiNamespace, sAxis := sSlave, sFb := 'GearIn',
       sMaster := sMaster, sTable := '', iParams := 5);
InGear := fbCall.InSync; Busy := fbCall.Busy; Active := fbCall.Active;
CommandAborted := fbCall.CommandAborted; Error := fbCall.Error; ErrorID := fbCall.ErrorID;
END_FUNCTION_BLOCK

FUNCTION_BLOCK SIM_MC_CamIn
VAR_INPUT
    Execute : BOOL; hConnection : DWORD; uiNamespace : UINT;
    sMaster : STRING(31); sSlave : STRING(31);
    MasterOffset : LREAL; SlaveOffset : LREAL; MasterScaling : LREAL := 1.0; SlaveScaling : LREAL := 1.0;
    StartMode : LREAL := 1.0;    (* 0 absolute, 1 relative *)
    CamTableID : LREAL;          (* 0 the table below, 1 the machine's own cam *)
    sTable : STRING(255);        (* lines 'master span, slave rise, law' or 'master, slave[, slope]' *)
END_VAR
VAR_OUTPUT
    InSync : BOOL; Busy : BOOL; Active : BOOL; CommandAborted : BOOL; Error : BOOL; ErrorID : UINT;
END_VAR
VAR
    fbCall : SIM_SyncHandshake;
END_VAR
fbCall.asParam[1] := 'MasterOffset';  fbCall.alrParam[1] := MasterOffset;
fbCall.asParam[2] := 'SlaveOffset';   fbCall.alrParam[2] := SlaveOffset;
fbCall.asParam[3] := 'MasterScaling'; fbCall.alrParam[3] := MasterScaling;
fbCall.asParam[4] := 'SlaveScaling';  fbCall.alrParam[4] := SlaveScaling;
fbCall.asParam[5] := 'StartMode';     fbCall.alrParam[5] := StartMode;
fbCall.asParam[6] := 'CamTableID';    fbCall.alrParam[6] := CamTableID;
fbCall(Execute := Execute, hConnection := hConnection, uiNamespace := uiNamespace, sAxis := sSlave, sFb := 'CamIn',
       sMaster := sMaster, sTable := sTable, iParams := 6);
InSync := fbCall.InSync; Busy := fbCall.Busy; Active := fbCall.Active;
CommandAborted := fbCall.CommandAborted; Error := fbCall.Error; ErrorID := fbCall.ErrorID;
END_FUNCTION_BLOCK

FUNCTION_BLOCK SIM_MC_GearOut
VAR_INPUT
    Execute : BOOL; hConnection : DWORD; uiNamespace : UINT; sSlave : STRING(31);
END_VAR
VAR_OUTPUT
    Done : BOOL; Busy : BOOL; Error : BOOL; ErrorID : UINT;
END_VAR
VAR
    fbCall : SIM_Handshake;
END_VAR
fbCall(Execute := Execute, hConnection := hConnection, uiNamespace := uiNamespace, sAxis := sSlave, sFb := 'GearOut', iParams := 0);
Done := fbCall.Done; Busy := fbCall.Busy; Error := fbCall.Error; ErrorID := fbCall.ErrorID;
END_FUNCTION_BLOCK

FUNCTION_BLOCK SIM_MC_CamOut
VAR_INPUT
    Execute : BOOL; hConnection : DWORD; uiNamespace : UINT; sSlave : STRING(31);
END_VAR
VAR_OUTPUT
    Done : BOOL; Busy : BOOL; Error : BOOL; ErrorID : UINT;
END_VAR
VAR
    fbCall : SIM_Handshake;
END_VAR
fbCall(Execute := Execute, hConnection := hConnection, uiNamespace := uiNamespace, sAxis := sSlave, sFb := 'CamOut', iParams := 0);
Done := fbCall.Done; Busy := fbCall.Busy; Error := fbCall.Error; ErrorID := fbCall.ErrorID;
END_FUNCTION_BLOCK

PROGRAM PRG_SimSyncDemo
VAR
    fbConnect    : UA_Connect;
    fbNamespace  : UA_NamespaceGetIndex;
    fbDisconnect : UA_Disconnect;
    stSession    : UASessionConnectInfo;
    hConnection  : DWORD;
    uiNamespace  : UINT;
    fbPowerX     : SIM_MC_Power;
    fbPowerY     : SIM_MC_Power;
    fbMoveX      : SIM_MC_MoveAbsolute;
    fbGearIn     : SIM_MC_GearIn;
    fbGearOut    : SIM_MC_GearOut;
    fbCamIn      : SIM_MC_CamIn;
    fbCamOut     : SIM_MC_CamOut;
    fbStopY      : SIM_MC_Stop;
    tonGeared    : TON;
    iStep        : INT;
    sMaster      : STRING(31) := 'x';    (* axis ids of the simulated machine: a two-axis gantry *)
    sSlave       : STRING(31) := 'y';
END_VAR

CASE iStep OF
0:  stSession.ApplicationName := 'CODESYS sim client';
    stSession.SecurityMsgMode := UASecurityMsgMode.UASMM_None;
    stSession.SecurityPolicy := UASecurityPolicy.UASP_None;
    fbConnect(Execute := TRUE, ServerEndpointUrl := 'opc.tcp://192.168.0.10:4840', SessionConnectInfo := stSession, Timeout := T#5S);
    IF fbConnect.Done THEN hConnection := fbConnect.ConnectionHdl; fbConnect(Execute := FALSE); iStep := 10;
    ELSIF fbConnect.Error THEN fbConnect(Execute := FALSE); iStep := 900; END_IF
10: fbNamespace(Execute := TRUE, ConnectionHdl := hConnection, NamespaceUri := 'urn:kinematics-simulation', Timeout := T#5S);
    IF fbNamespace.Done THEN uiNamespace := fbNamespace.NamespaceIndex; fbNamespace(Execute := FALSE); iStep := 20;
    ELSIF fbNamespace.Error THEN fbNamespace(Execute := FALSE); iStep := 900; END_IF
20: fbPowerX.Enable := TRUE; fbPowerY.Enable := TRUE;
    IF fbPowerX.Status AND fbPowerY.Status THEN iStep := 30; END_IF
30: (* the master runs slowly over its stroke *)
    fbMoveX.Position := 0.9; fbMoveX.Velocity := 0.05; fbMoveX.Acceleration := 1.0; fbMoveX.Deceleration := 1.0;
    fbMoveX.Jerk := 100.0; fbMoveX.Execute := TRUE;
    IF fbMoveX.Busy THEN iStep := 40; ELSIF fbMoveX.Error THEN iStep := 900; END_IF
40: (* y gears in at 2:1 *)
    fbGearIn.RatioNumerator := 2.0; fbGearIn.RatioDenominator := 1.0;
    fbGearIn.Acceleration := 1.0; fbGearIn.Deceleration := 1.0; fbGearIn.Jerk := 100.0;
    fbGearIn.Execute := TRUE;
    tonGeared(IN := fbGearIn.InGear, PT := T#1S);
    IF tonGeared.Q THEN iStep := 50; ELSIF fbGearIn.Error OR fbGearIn.CommandAborted THEN iStep := 900; END_IF
50: fbGearOut.Execute := TRUE;
    IF fbGearOut.Done THEN fbGearOut.Execute := FALSE; fbGearIn.Execute := FALSE; iStep := 60;
    ELSIF fbGearOut.Error THEN iStep := 900; END_IF
60: (* y cams in, relative, on a 3-4-5 rise of 20 mm over 0.1 m of x and back *)
    fbCamIn.sTable := '0.1, 0.02, 3-4-5$N0.1, -0.02, 3-4-5';
    fbCamIn.StartMode := 1.0; fbCamIn.CamTableID := 0.0;
    fbCamIn.Execute := TRUE;
    IF fbCamIn.InSync THEN iStep := 70; ELSIF fbCamIn.Error THEN iStep := 900; END_IF
70: IF NOT fbMoveX.Busy THEN iStep := 80; END_IF   (* x has arrived; y stands on its cam *)
80: fbCamOut.Execute := TRUE;
    IF fbCamOut.Done THEN fbCamOut.Execute := FALSE; fbCamIn.Execute := FALSE; iStep := 90;
    ELSIF fbCamOut.Error THEN iStep := 900; END_IF
90: fbStopY.Deceleration := 1.0; fbStopY.Execute := TRUE;
    IF fbStopY.Done THEN fbStopY.Execute := FALSE; fbMoveX.Execute := FALSE; iStep := 95;
    ELSIF fbStopY.Error THEN iStep := 900; END_IF
95: fbPowerX.Enable := FALSE; fbPowerY.Enable := FALSE;
    IF NOT fbPowerX.Status AND NOT fbPowerY.Status THEN iStep := 99; END_IF
99: fbDisconnect(Execute := TRUE, ConnectionHdl := hConnection, Timeout := T#5S);
    IF fbDisconnect.Done OR fbDisconnect.Error THEN fbDisconnect(Execute := FALSE); iStep := 100; END_IF
100: ;
900: ;
END_CASE

IF iStep >= 20 AND iStep < 99 THEN
    fbPowerX(hConnection := hConnection, uiNamespace := uiNamespace, sAxis := sMaster);
    fbPowerY(hConnection := hConnection, uiNamespace := uiNamespace, sAxis := sSlave);
    fbMoveX(hConnection := hConnection, uiNamespace := uiNamespace, sAxis := sMaster);
    fbGearIn(hConnection := hConnection, uiNamespace := uiNamespace, sMaster := sMaster, sSlave := sSlave);
    fbGearOut(hConnection := hConnection, uiNamespace := uiNamespace, sSlave := sSlave);
    fbCamIn(hConnection := hConnection, uiNamespace := uiNamespace, sMaster := sMaster, sSlave := sSlave);
    fbCamOut(hConnection := hConnection, uiNamespace := uiNamespace, sSlave := sSlave);
    fbStopY(hConnection := hConnection, uiNamespace := uiNamespace, sAxis := sSlave);
END_IF
END_PROGRAM
